Fanuc KAREL source: KC00041.KL

PROGRAM KC00041
%NOLOCKGROUP
%ENVIRONMENT IOSETUP
VAR
  I: INTEGER
  J: INTEGER
  K: INTEGER
  R: REAL
  B: BOOLEAN
  S: STRING[80]
  T: STRING[80]
  P: PATH
  Q: PATH
  AI: ARRAY[8] OF INTEGER
  AB: ARRAY[244] OF BYTE
BEGIN
  GET_PORT_VAL(I,J,K,I)
END KC00041
